Staubli VAL3: PrecProg.pjx

--- PrecProg.pjx ---
Parameters version=s7.5.3 stackSize=5000 millimeterUnit=true
Program file=MoveJoint.pgx
Program file=MoveLine.pgx
Program file=start.pgx
Program file=stop.pgx
Program file=main.pgx
Data file=PrecProg.dtx

--- PrecProg.dtx ---
mdesc mNomSpeed
frame fFrame1 = {x=0.000, y=-0.001, z=1000.000, rx=90.000, ry=0.123, rz=0.500, fatherId=world[0]}
dio Input[16]
  [0] = {link=BasicIO-1\%I0}
  [1] = {link=BasicIO-1\%I1}
  [2] = {link=BasicIO-1\%I2}
  [3] = {link=BasicIO-1\%I3}
  [4] = {link=BasicIO-1\%I4}
  [5] = {link=BasicIO-1\%I5}
  [6] = {link=BasicIO-1\%I6}
  [7] = {link=BasicIO-1\%I7}
  [8] = {link=BasicIO-1\%I8}
  [9] = {link=BasicIO-1\%I9}
  [10] = {link=BasicIO-1\%I10}
  [11] = {link=BasicIO-1\%I11}
  [12] = {link=BasicIO-1\%I12}
  [13] = {link=BasicIO-1\%I13}
  [14] = {link=BasicIO-1\%I14}
  [15] = {link=BasicIO-1\%I15}
dio Output[16]
  [0] = {link=BasicIO-1\%Q0}
  [1] = {link=BasicIO-1\%Q1}
  [2] = {link=BasicIO-1\%Q2}
  [3] = {link=BasicIO-1\%Q3}
  [4] = {link=BasicIO-1\%Q4}
  [5] = {link=BasicIO-1\%Q5}
  [6] = {link=BasicIO-1\%Q6}
  [7] = {link=BasicIO-1\%Q7}
  [8] = {link=BasicIO-1\%Q8}
  [9] = {link=BasicIO-1\%Q9}
  [10] = {link=BasicIO-1\%Q10}
  [11] = {link=BasicIO-1\%Q11}
  [12] = {link=BasicIO-1\%Q12}
  [13] = {link=BasicIO-1\%Q13}
  [14] = {link=BasicIO-1\%Q14}
  [15] = {link=BasicIO-1\%Q15}
tool tCurrentTool = {x=0.125, y=-0.375, z=123.457, rx=-45.250, ry=-0.000, rz=0.000, fatherId=flange[0], ioLink=ValveIO/valve1}
mdesc mCurrentSpeed
pointRs pPointRs = {fatherId=fFrame1[0]}
pointRs pPointRs2 = {fatherId=fFrame1[0]}

--- main.pgx ---
program main()
begin
  close(tCurrentTool)
  pPointRs.config.shoulder = lefty
  pPointRs2.config.shoulder = lefty
  mCurrentSpeed.tvel = 100.00
  mCurrentSpeed.blend = joint
  mCurrentSpeed.reach = 0.010
  mCurrentSpeed.leave = 0.010
  // Program PrecProg start
  // Program generated by RoboDK v6.0.7 for Staubli TS20 FL 100 TC on XX/XX/XXXX 18:00:00
  // Using nominal kinematics.
  call MoveJoint(12.34560,-45.67890,78.90130,-0.50000)
  call MoveLine(-640.585,506.981,371.534,136.641,31.137,-130.569)
  call MoveLine(0.500,-0.500,0.250,-180.000,0.005,-0.005)
  call MoveJoint(-12.34540,45.67850,-78.90000,0.50000)
  call MoveJoint(-12.34540,45.67850,-78.90000,0.50000)
  mCurrentSpeed.tvel = 66.667
  delay(0.002)
  delay(1.000)
  call MoveLine(-353.026,-90.135,331.702,164.619,39.324,-168.579)

  waitEndMove()
  // Program PrecProg end

end

--- start.pgx ---
program start()
begin
  call main()
end

--- MoveJoint.pgx ---
program MoveJoint(num x_nJ1, num x_nJ2, num x_nJ3, num x_nJ4)
  local joint l_jJoint
begin
  l_jJoint.j1 = x_nJ1
  l_jJoint.j2 = x_nJ2
  l_jJoint.j3 = x_nJ3
  l_jJoint.j4 = x_nJ4
  movej(l_jJoint,tCurrentTool ,mCurrentSpeed)
end

--- MoveLine.pgx ---
program MoveLine(num x_nX, num x_nY, num x_nZ, num x_nRx, num x_nRy, num x_nRz)
begin
  pPointRs.trsf.x = x_nX
  pPointRs.trsf.y = x_nY
  pPointRs.trsf.z = x_nZ
  pPointRs.trsf.rx = x_nRx
  pPointRs.trsf.ry = x_nRy
  pPointRs.trsf.rz = x_nRz
  movel(pPointRs,tCurrentTool,mCurrentSpeed)
end

--- stop.pgx ---
program stop()
begin
end
